// TIA Portal V18 export
VAR_GLOBAL   // PLC tag table "BYPASS_STATIONS"
   BYPASS_STATION_1 AT %M36.2 : Bool;
   BYPASS_POSTO_1 AT %M36.3 : Bool;
   BYPASS_STATION_5 AT %M36.4 : Bool;
   BYPASS_POSTO_5 AT %M36.5 : Bool;
   BYPASS_STATION_10 AT %M36.6 : Bool;
   BYPASS_POSTO_10 AT %M36.7 : Bool;
   BYPASS_STATION_15 AT %M37.0 : Bool;
   BYPASS_POSTO_15 AT %M37.1 : Bool;
   BYPASS_STATION_20 AT %M37.2 : Bool;
   BYPASS_POSTO_20 AT %M37.3 : Bool;
   BYPASS_STATION_30 AT %M37.4 : Bool;
   BYPASS_POSTO_30 AT %M37.5 : Bool;
   BYPASS_STATION_40 AT %M37.6 : Bool;
   BYPASS_POSTO_40 AT %M37.7 : Bool;
   BYPASS_STATION_50 AT %M38.0 : Bool;
   BYPASS_POSTO_50 AT %M38.1 : Bool;
   BYPASS_STATION_55 AT %M38.2 : Bool;
   BYPASS_POSTO_55 AT %M38.3 : Bool;
   BYPASS_STATION_60 AT %M38.4 : Bool;
   BYPASS_POSTO_60 AT %M38.5 : Bool;
   BYPASS_STATION_70 AT %M38.6 : Bool;
   BYPASS_POSTO_70 AT %M38.7 : Bool;
   BYPASS_STATION_75 AT %M39.0 : Bool;
   BYPASS_POSTO_75 AT %M39.1 : Bool;
   BYPASS_STATION_80 AT %M39.2 : Bool;
   BYPASS_POSTO_80 AT %M39.3 : Bool;
   BYPASS_STATION_90 AT %M39.4 : Bool;
   BYPASS_POSTO_90 AT %M39.5 : Bool;
   BYPASS_STATION_95 AT %M39.6 : Bool;
   BYPASS_POSTO_95 AT %M39.7 : Bool;
   BYPASS_STATION_100 AT %M40.0 : Bool;
   BYPASS_POSTO_100 AT %M40.1 : Bool;
   BYPASS_STATION_105 AT %M40.2 : Bool;
   BYPASS_POSTO_105 AT %M40.3 : Bool;
   BYPASS_STATION_110 AT %M40.4 : Bool;
   BYPASS_POSTO_110 AT %M40.5 : Bool;
   BYPASS_STATION_115 AT %M40.6 : Bool;
   BYPASS_POSTO_115 AT %M40.7 : Bool;
   BYPASS_STATION_120 AT %M41.0 : Bool;
   BYPASS_POSTO_120 AT %M41.1 : Bool;
   BYPASS_STATION_125 AT %M41.2 : Bool;
   BYPASS_POSTO_125 AT %M41.3 : Bool;
   BYPASS_STATION_130 AT %M41.4 : Bool;
   BYPASS_POSTO_130 AT %M41.5 : Bool;
   BYPASS_STATION_140 AT %M41.6 : Bool;
   BYPASS_POSTO_140 AT %M41.7 : Bool;
   BYPASS_STATION_150 AT %M42.0 : Bool;
   BYPASS_POSTO_150 AT %M42.1 : Bool;
   BYPASS_STATION_QG AT %M42.2 : Bool;
   BYPASS_POSTO_QG AT %M42.3 : Bool;
END_VAR
